FUNCTION_BLOCK ABSTRACT FB_Device
VAR_OUTPUT
	bFault : BOOL;   // device fault
END_VAR

END_FUNCTION_BLOCK

(* stored: Version 1.1.0.1, ProductVersion 3.1.4026.12
   POU FB_Device: Id {3a2b3c4d-0000-4000-8000-000000000005}, SpecialFunc None *)
